// TIA Portal V21 export
// export: Created 2026-08-21T20:18:54.5743067Z, ExportSetting None, DisplayName Totally Integrated Automation Portal, DisplayVersion V21, DisplayName STEP 7 Professional, DisplayVersion V21, DisplayName STEP 7 Safety, DisplayVersion V21, DisplayName Tech WebApplication, DisplayVersion V21, DisplayName WinCC Basic/Comfort/Advanced, DisplayVersion V21, DisplayName WinCC Professional, DisplayVersion V21, DisplayName WinCC Unified, DisplayVersion V21
TYPE "UDT_MTP_BinReportValue"
   STRUCT
      WQC { ExternalWritable := 'False'} : Byte := 16#FF;   // Worst Quality Code
      V { ExternalWritable := 'False'} : Bool;   // Value
      VState0 { ExternalWritable := 'False'} : String[16];   // text replacement for false
      VState1 { ExternalWritable := 'False'} : String[16];   // text replacement for true
      MissedValue { ExternalWritable := 'False'} : Bool;   // MissedValueFeature
   END_STRUCT;
END_TYPE
